    PGN_PROPRIETARY_B_PAGE_1_131042 : UDINT := UDINT#16#1FFE2; (* < 131042 - PropB1_E2 *)
    PGN_PROPRIETARY_B_PAGE_1_131043 : UDINT := UDINT#16#1FFE3; (* < 131043 - PropB1_E3 *)
    PGN_PROPRIETARY_B_PAGE_1_131044 : UDINT := UDINT#16#1FFE4; (* < 131044 - PropB1_E4 *)
    PGN_PROPRIETARY_B_PAGE_1_131045 : UDINT := UDINT#16#1FFE5; (* < 131045 - PropB1_E5 *)
    PGN_PROPRIETARY_B_PAGE_1_131046 : UDINT := UDINT#16#1FFE6; (* < 131046 - PropB1_E6 *)
    PGN_PROPRIETARY_B_PAGE_1_131047 : UDINT := UDINT#16#1FFE7; (* < 131047 - PropB1_E7 *)
    PGN_PROPRIETARY_B_PAGE_1_131048 : UDINT := UDINT#16#1FFE8; (* < 131048 - PropB1_E8 *)
    PGN_PROPRIETARY_B_PAGE_1_131049 : UDINT := UDINT#16#1FFE9; (* < 131049 - PropB1_E9 *)
    PGN_PROPRIETARY_B_PAGE_1_131050 : UDINT := UDINT#16#1FFEA; (* < 131050 - PropB1_EA *)
    PGN_PROPRIETARY_B_PAGE_1_131051 : UDINT := UDINT#16#1FFEB; (* < 131051 - PropB1_EB *)
    PGN_PROPRIETARY_B_PAGE_1_131052 : UDINT := UDINT#16#1FFEC; (* < 131052 - PropB1_EC *)
    PGN_PROPRIETARY_B_PAGE_1_131053 : UDINT := UDINT#16#1FFED; (* < 131053 - PropB1_ED *)
    PGN_PROPRIETARY_B_PAGE_1_131054 : UDINT := UDINT#16#1FFEE; (* < 131054 - PropB1_EE *)
    PGN_PROPRIETARY_B_PAGE_1_131055 : UDINT := UDINT#16#1FFEF; (* < 131055 - PropB1_EF *)
    PGN_PROPRIETARY_B_PAGE_1_131056 : UDINT := UDINT#16#1FFF0; (* < 131056 - PropB1_F0 *)
    PGN_PROPRIETARY_B_PAGE_1_131057 : UDINT := UDINT#16#1FFF1; (* < 131057 - PropB1_F1 *)
    PGN_PROPRIETARY_B_PAGE_1_131058 : UDINT := UDINT#16#1FFF2; (* < 131058 - PropB1_F2 *)
    PGN_PROPRIETARY_B_PAGE_1_131059 : UDINT := UDINT#16#1FFF3; (* < 131059 - PropB1_F3 *)
    PGN_PROPRIETARY_B_PAGE_1_131060 : UDINT := UDINT#16#1FFF4; (* < 131060 - PropB1_F4 *)
    PGN_PROPRIETARY_B_PAGE_1_131061 : UDINT := UDINT#16#1FFF5; (* < 131061 - PropB1_F5 *)
    PGN_PROPRIETARY_B_PAGE_1_131062 : UDINT := UDINT#16#1FFF6; (* < 131062 - PropB1_F6 *)
    PGN_PROPRIETARY_B_PAGE_1_131063 : UDINT := UDINT#16#1FFF7; (* < 131063 - PropB1_F7 *)
    PGN_PROPRIETARY_B_PAGE_1_131064 : UDINT := UDINT#16#1FFF8; (* < 131064 - PropB1_F8 *)
    PGN_PROPRIETARY_B_PAGE_1_131065 : UDINT := UDINT#16#1FFF9; (* < 131065 - PropB1_F9 *)
    PGN_PROPRIETARY_B_PAGE_1_131066 : UDINT := UDINT#16#1FFFA; (* < 131066 - PropB1_FA *)
    PGN_PROPRIETARY_B_PAGE_1_131067 : UDINT := UDINT#16#1FFFB; (* < 131067 - PropB1_FB *)
    PGN_PROPRIETARY_B_PAGE_1_131068 : UDINT := UDINT#16#1FFFC; (* < 131068 - PropB1_FC *)
    PGN_PROPRIETARY_B_PAGE_1_131069 : UDINT := UDINT#16#1FFFD; (* < 131069 - PropB1_FD *)
    PGN_PROPRIETARY_B_PAGE_1_131070 : UDINT := UDINT#16#1FFFE; (* < 131070 - PropB1_FE *)
    PGN_PROPRIETARY_B_PAGE_1_LAST_ENTRY : UDINT := UDINT#16#1FFFF; (* < 131071 - PropB1_FF *)
  END_VAR
END_GLOBALCONSTANTS
